(* IEC 61131-3 sources: kns-port-domestic/tools/port_metrics_tests/fixtures/adapted/src/POUs/FB_VfdLink_Regul, 1 file *)

(* ---- FB_VfdLink_Regul.decl.st ---- *)
// PORT: адаптер связи с ПЧ через Modbus Serial Master вместо устройства CODESYS
FUNCTION_BLOCK FB_VfdLink_Regul
VAR_INPUT
    awData : ARRAY[0..3] OF WORD;
END_VAR
VAR_OUTPUT
    rSpeed_Hz : REAL;
END_VAR
